Universal Robots URScript: T002_zai-org_GLM-4.7-FP8_edit_perf_rep1.urscript

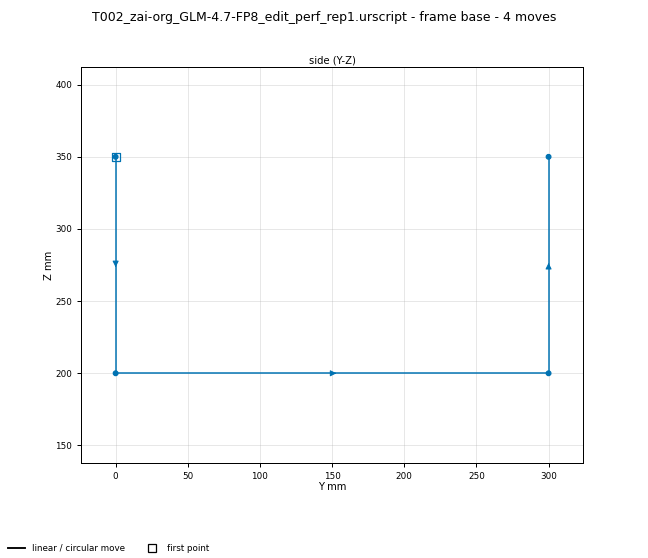
[picture p0: tool path of T002_zai-org_GLM-4.7-FP8_edit_perf_rep1.urscript in frame base, 4 of 6 moves have a stored position in this frame; points joined in program order, loops and branches not executed]
# Task: T002 — Linear weld path — fenced mode (Optimized)
# Generated by ENFIELD IR→URScript Translator
# Operating mode: fenced | Max TCP speed: 0.500 m/s
# Robot: ur5e
#
# WARNING: This is auto-generated code for SIMULATION ONLY.
# Do NOT deploy to a physical robot without safety review.

def task_T002():
  # [0] Verify E-Stop clear before weld sequence
  if (get_digital_in(0) == True):
    popup("E-Stop active — aborting program.", error=True)
    halt
  end

  # [Optimization] Start Gas Pre-flow early to overlap with motion
  set_digital_out(1, True)

  # [1] Go to home position (Increased velocity/acceleration)
  movej([0.0000, -1.5708, 1.5708, -1.5708, -1.5708, 0.0000], a=2.0000, v=1.5000)

  # [2] Approach above weld start (Max TCP speed, increased blend radius)
  movel(p[0.450000, 0.000000, 0.350000, 0.0000, 3.1416, 0.0000], a=1.2000, v=0.5000, r=0.0500)

  # [3] Descend to weld start position (Faster approach, precise stop)
  # Gas pre-flow delay (0.5s) is covered by the motion time from Home
  movel(p[0.450000, 0.000000, 0.200000, 0.0000, 3.1416, 0.0000], a=0.5000, v=0.3000, r=0.0000)

  # [4] Arc ON — welding start
  set_digital_out(0, True)
  set_analog_out(0, 0.400)
  set_analog_out(1, 0.333)

  # [5] Weld seam — 300mm linear path (Process speed maintained, accel increased)
  movel(p[0.450000, 0.300000, 0.200000, 0.0000, 3.1416, 0.0000], a=0.5000, v=0.0500)

  # [6] Arc OFF — welding end
  set_digital_out(0, False)
  set_analog_out(0, 0.0)
  set_analog_out(1, 0.0)

  # [7] Retract above weld end (Max speed, overlapping with post-flow delay)
  movel(p[0.450000, 0.300000, 0.350000, 0.0000, 3.1416, 0.0000], a=1.2000, v=0.5000, r=0.0500)

  # [8] Post-weld gas flow (Delay occurs after retract is complete)
  sleep(1.0000)

  # [9] Gas flow OFF
  set_digital_out(1, False)

  # [10] Return to home (Increased velocity/acceleration)
  movej([0.0000, -1.5708, 1.5708, -1.5708, -1.5708, 0.0000], a=2.0000, v=1.5000)

end

# Entry point
task_T002()
